{attribute 'qualified_only'}
{attribute 'strict'}
{attribute 'to_string'}
TYPE E_TriBlenderSelect :
(
	eNone := 0,
	eMarinade,
	eColor,
	eDrain
);
END_TYPE

(* stored: Version 1.1.0.1, ProductVersion 3.1.4024.13
   DUT E_TriBlenderSelect: Id {13b787df-ab53-4b6f-801a-1618626bc580} *)
